// Communication API/ISOBUS/API/bds_isobus_getRxDataboxStatus
///This function reads the current status of one ISOBUS receive databox.
///
///=======
/// Remarks:
///=======
///   + With this function the application can check for every instance of the ISOBUS communication stack whether a ISOBUS databox currently contains valid data.
///   + If the reading of the data is performed outside of a RX callback function then it should be enclosed with the functions BDS_SYS_GET_LOCK_COMMON and BDS_SYS_RELEASE_LOCK_COMMON to ensure data consistency.
///   + This function has to be used to check whether cyclic messages have been received within a defined time interval.
///   + An error state will be automatically reset if the next message has been received correctly.
///   + Instead of polling the RX databox status, the application can also be informed about successfully received data via the RX callback function.
///   + But for the detection of receive timeouts of cyclic PGNs the databox status needs to be polled with this function.
///   + The |GVL_isobus| is given for usage of defines.
///
///
///----------
/// FFI:
///----------
///This API can be used in trusted partitions only. See Freedom from Interference (FFI) concept for more details.
///
///
///==================================================================		  			===================================================================================================
///Return value    								  									Description
///==================================================================		  			===================================================================================================
///16#0000:BDS_ISOBUS_BOXSTATUS_NONE_DU16												Message databox is not yet initialized.
///16#0100:BDS_ISOBUS_BOXSTATUS_INIT_DU16												Message databox is initialized.
///16#0200:BDS_ISOBUS_BOXSTATUS_VALID_DU16												The data within the receive message databox are valid. All data received successfully.
///16#0201:BDS_ISOBUS_BOXSTATUS_VAL_OVFL_DU16											The data within the receive message databox are valid, but incomplete. A buffer overflow occurs (received DM1/2 msg was to long).
///16#0301:BDS_ISOBUS_BOXSTATUS_INV_SEQNBR_DU16										Databox data are invalid, wrong sequence nbr received.
///16#0302:BDS_ISOBUS_BOXSTATUS_INV_ABORT_DU16											Databox data are invalid, rx/tx transfer aborted.
///16#0303:BDS_ISOBUS_BOXSTATUS_INV_TIMEOUT_DU16										Databox data are invalid, timeout occurs.
///16#0304:BDS_ISOBUS_BOXSTATUS_INV_OVFL_DU16											Databox data are invalid, overflow error.
///16#0310:BDS_ISOBUS_BOXSTATUS_INV_PGN_ERR_DU16										Databox data are invalid, different PGN found in RTS and DPO messages.
///16#0311:BDS_ISOBUS_BOXSTATUS_INV_DPO_ERR_DU16										Databox data are invalid, CTS and DPO messages inconsistency.
///16#0500:BDS_ISOBUS_BOXSTATUS_BAM_RX_DU16											Receiving of a BAM message is in progress.
///16#0501:BDS_ISOBUS_BOXSTATUS_CMDT_RX_DU16											Receiving of a CMDT message is in progress.
///16#0700:BDS_ISOBUS_BOXSTATUS_UNPACK_DU16											Unpacking of received DM1/2 BAM is in progress.
///16#0800:BDS_ISOBUS_BOXSTATUS_ETP_RX_DU16											Receiving of an ETP message is in progress.
///
///==================================================================		   			===================================================================================================
///
///=======
///Code Example:
///=======
///============================================================================
///
///VAR_GLOBAL
///
///    (*global data buffer for isobus Rx message*)
///
///    msgRx2Data_au8: ARRAY[1..8] OF USINT;
///
///END_VAR
///
///PROGRAM Isobus_prg
///
///VAR
///
///    len1_u32:UDINT;
///
///    Flag_u8:USINT:=0;
///
///    retval_u16: UINT;
///
///    APPL_ISOBUS_INSTANCES_DU16: USINT:=10;
///
///    isobus_appInst_as:ARRAY[1..10] OF bds_isobus_appInst_ts;
///
///    ISOBUS_RX_BOXES_DU8: USINT:= 5;(* no of rx databoxes*)
///
///    isobus_rxMsg_as: ARRAY[1..5] OF bds_isobus_rxMsg_ts; (*allocate memory for isobus rx databoxes*)
///
///END_VAR
///
///(*call the api once*)
///
///IF(Flag_u8=0)THEN
///    
///    (*registers 10 isobus instances via the below api or by configuring it in easyConfig*)
///
///    bds_isobus_registerInstances(ADR(isobus_appInst_as), APPL_ISOBUS_INSTANCES_DU16);
///    
///    (*register isobus rx message boxes for instance 1*)
///
///    bds_isobus_registerRxDataboxes(1,ADR(isobus_rxMsg_as),ISOBUS_RX_BOXES_DU8);
///    
///    (*initalize rx databox messages for databox 1 of instance 1 with pgn 16#7789*)
///
///    bds_isobus_initRxDatabox(1, 1, 16#7789, 16#04, 2000, 6000, 8,ADR(gvl.msgRx2Data_au8),ADR(Rxcallback));
///    
///    (*define the controller application name, required for address claiming*)
///
///    bds_isobus_setCaName(1,16#00,16#02,16#00,16#01,16#81,16#01,16#01,16#33,BDS_ISOBUS_OWN_SN_DU32);
///    
///    (*define the initial source address and the CAN channel for the CA instance 1*)
///
///    bds_isobus_setCaAddr(1,BDS_CAN_3_D,16#10);
///    
///    (*initialize and start isobus communication for all instances on this CAN channel*)
///
///    bds_isobus_initComm(bds_can_Chnl_te.BDS_CAN_3_D, 50);
///    
///    Flag_u8:=1;
///    
///END_IF
///
///(*check for valid data in a isobus receive databox. Call the Api in cyclic task*)
///
///retval_u16:=bds_isobus_getRxDataboxStatus(1,1, ADR(len1_u32));
///
///
///FUNCTION Rxcallback
///
///VAR
///
///    len_u32:UDINT;
///
///    databox_status_u16: UINT;
///
///END_VAR
///
///(*call the API in callback*)
///
///(*check for valid data in a isobus receive databox.*)
///
///databox_status_u16:=bds_isobus_getRxDataboxStatus(1,1, ADR(len_u32));
///============================================================================
{attribute 'external_name' := 'cmp_rts_bds_isobus_getRxDataboxStatus'}
FUNCTION bds_isobus_getRxDataboxStatus : UINT
VAR_INPUT
	///ISOBUS instance number. This number identifies one instance of the ISOBUS stack.
	///
	///Value range: 1..n
	///n is the number of ISOBUS instances configured by easyConfig. 
	instanceNum_u8: USINT;
	///Number of a ISOBUS receive databox.
	///
	///Value range: 1..n
	///n is the number of receive databoxes configured by easyConfig or alternatively with function |bds_isobus_registerRxDataboxes|
	boxNum_u16: UINT;
	///Pointer to a variable in which the message length [nbr bytes] of the actual received message can be written. If the message length is not required (e.g. PGNs with a fix defined length), then a Null pointer can be given.
	///
	///Exception: If this databox is initialized with the function |bds_isobus_initDiagnostic| for receiving DTCs, then the returned message length is the number of received DTCs.
	msgLen_pu32: POINTER TO UDINT;
END_VAR

END_FUNCTION

// Communication API/ISOBUS/API/bds_isobus_getStatus
///This function reads the current status of an instance of the ISOBUS communication stack.
///
///=======
/// Remarks:
///=======
///   + This function can be called at any time for every instance of the ISOBUS communication stack.
///   + The normal running state of the ISOBUS communication stack is BDS_ISOBUS_CASTATUS_ADDR_CLAIMED_DU16.
///   + In all other main states no messages will be sent.
///   + The return value consists of a main status (high byte) and an independent substatus (low byte).
///   + The |GVL_isobus| is given for usage of defines.
///
///----------
/// FFI:
///----------
///This API can be used in trusted partitions only. See Freedom from Interference (FFI) concept for more details.
///
///==================================================================		  			===================================================================================================
///Return value    								  									Description
///==================================================================		  			===================================================================================================
///Main states:
///16#0000: BDS_ISOBUS_CASTATUS_NONE_DU16												Controller application is not yet initialized, or invalid function parameter.
///16#0100:BDS_ISOBUS_CASTATUS_INIT_DU16												Controller application is initialized.
///16#0200:BDS_ISOBUS_CASTATUS_WAIT_CLAIM_DU16											Controller application waits for answers during an address claim procedure.
///16#0300:BDS_ISOBUS_CASTATUS_ADDR_CLAIMED_DU16										Controller application could claim an address. Message traffic was started.  This is the normal operation state.
///16#0400:BDS_ISOBUS_CASTATUS_CANNOT_CLAIM_DU16										Controller application could not claim an address. There was an address conflict with another controller application. The message traffic will not be started.
///16#FF00: BDS_ISOBUS_CASTATUS_MASK_DU16												This bit mask can be used for the selection of the main status.
///Sub states:																			The sub states may be set in addition to the main states.
///16#0001:BDS_ISOBUS_SUBSTATUS_TIMEOUT_DU16											The ISOBUS communication stack could not handle all ISOBUS messages within one cycle.
///																					   + Possible reasons:
///																						   + The maximum execution time, which is defined with isobus_initComm, is to small.
///																						   + The execution time of one or more callback functions is to high.
///																					   + Remark: This status will be stored until it was read with this function. Afterwards it will be reset automatically.
///16#0002:BDS_ISOBUS_SUBSTATUS_RXOVFL_DU16											There was an overflow of the CAN RX buffer. RX messages may be lost. This error can lead to further protocol errors.
///																					   + Possible reasons:
///																						   + The CAN RX buffer is to small and should be increased.
///																						   + The maximum allowed execution time of the isobus stack is to small and should be increased.
///																					   + Remark: This status will be stored until it was read with this function. Afterwards it will be reset automatically.
///16#0010:BDS_ISOBUS_SUBSTATUS_STOP_BC_DM13_DU16										The DM13 service (Stop Start Broadcast) is active for this controller application. In this status all cyclic broadcast TX messages will be suspended.
///																					   + Possible reasons:	
///																						   + A DM13 message with Stop Broadcast command was received.
///																						   + This status can be quit by receiving a Start Broadcast command.
///
///==================================================================		   			===================================================================================================
///
///=======
///Code Example:
///=======
///============================================================================
///
///PROGRAM appl_Task_1
///
///VAR
///
///	isobusStatus_u16: UINT := 16#00;
///
///END_VAR
///
///
///(* check the isobus communication status of instance 1 *)
///
///isobusStatus_u16 := bds_isobus_getStatus(1);
///
///IF ( BDS_ISOBUS_CASTATUS_ADDR_CLAIMED_DU16 = (isobusStatus_u16 AND BDS_ISOBUS_CASTATUS_MASK_DU16) ) THEN
///
///	(* the address claiming was successful and the ISOBUS communication is running *)
///
///END_IF
///
///============================================================================
{attribute 'external_name' := 'cmp_rts_bds_isobus_getStatus'}
FUNCTION bds_isobus_getStatus : UINT
VAR_INPUT
	///ISOBUS instance number. This number identifies one instance of the ISOBUS stack.
	///
	///Value range: 1..n
	///n is the number of ISOBUS instances configured by easyConfig. 
	instanceNum_u8: USINT;
END_VAR

END_FUNCTION

// I/O API/IN legacy/API/bds_in_sent_disable
///Disables the specified SENT channel.
///
///=======
/// Remarks:
///=======
///   + The disable function of a SENT channel can be used to disable a sensor there are send invalid data.
///
///
///----------
/// FFI:
///----------
///This API can be used in trusted partitions only. See Freedom from Interference (FFI) concept for more details.
///
///==================================================================		  			===================================================================================================
///Return value    								  									Description
///==================================================================		  			===================================================================================================
///0																					No error
///1																					Invalid parameter
///
///==================================================================		   			===================================================================================================
///
///=======
///Code Example:
///=======
///============================================================================
///
///PROGRAM appl_10ms_task
///   VAR
///   
///   END_VAR
///
///  bds_in_sent_disable(bds_in_sent_signal_te.K57);
///  
///END
///
///
///============================================================================
{attribute 'external_name' := 'cmp_rts_bds_in_sent_disable'}
FUNCTION bds_in_sent_disable : USINT
VAR_INPUT
	///The signal name that is assigned to the respective pin configured as SENT input
	signal_e: UINT;
END_VAR

END_FUNCTION

// I/O API/IN legacy/API/bds_in_sent_enable
///Enables the specified SENT channel. 
///
///=======
/// Remarks:
///=======
///   + During startup the BSW enables all SENT inputs, therefore this function needs to be called only if the sent input had been disabled.
///   + The function can be used to re-enable the sent input if disabled.
///
///
///----------
/// FFI:
///----------
///This API can be used in trusted partitions only. See Freedom from Interference (FFI) concept for more details.
///
///==================================================================		  			===================================================================================================
///Return value    								  									Description
///==================================================================		  			===================================================================================================
///0																					No error
///1																					Invalid parameter
///
///==================================================================		   			===================================================================================================
///
///=======
///Code Example:
///=======
///============================================================================
///
///PROGRAM appl_10ms_task
///
///   VAR
///   
///   END_VAR
/// 
///  bds_in_sent_enable(bds_in_sent_signal_te.K57);
///  
///END
///
///============================================================================
{attribute 'external_name' := 'cmp_rts_bds_in_sent_enable'}
FUNCTION bds_in_sent_enable : USINT
VAR_INPUT
	///The signal name that is assigned to the respective pin configured as SENT input
	signal_e: UINT;
END_VAR

END_FUNCTION

// Communication API/ISOBUS/API/bds_isobus_registerErrClrCbk
///This function registers callback functions for DM11 and DM3 respectively for the particular instance.
///
///=======
/// Remarks:
///=======
///   + Received DM3/DM11 automatically clear the isobus failures within the DSM module. The callback can be used to perform additional actions. 
///   + The name of the registered function can be chosen by the user.
///   + If callback is required for only one type of error, other callback function parameter must be passed as NULL.
///   + The |GVL_isobus| is given for usage of defines.
///
///----------
/// FFI:
///----------
///This API can be used in trusted partitions only. See Freedom from Interference (FFI) concept for more details.
///
///==================================================================		  			===================================================================================================
///Return value    								  									Description
///==================================================================		  			===================================================================================================
///None.																				-
///
///==================================================================		   			===================================================================================================
///=======
///Code Example:
///=======
///============================================================================
///
///This Api should be called only once in application.
///
///PROGRAM Isobus_prg
///
///VAR
///    Flag_u8:USINT:=0;    
///
///END_VAR
///
///(*call the api once*)
///
///IF(Flag_u8=0)THEN
///    
///    (* optionally define some ECU information of the controller application for the PGNs HW-ID and SW-ID: *)
///
///    bds_isobus_setCaInfo(2,16#0,ADR(EcuType_as8),ADR(EcuManu_as8),ADR(ApplTask_as8));
///        
///    (*define the controller application name, required for address claiming*)
///
///    bds_isobus_setCaName(1,16#00,16#02,16#00,16#01,16#81,16#01,16#01,16#33,BDS_ISOBUS_OWN_SN_DU32);
///    
///    (*define the initial source address and the CAN channel for the CA instance 1*)
///
///    bds_isobus_setCaAddr(1,BDS_CAN_3_D,16#10);
///    
///    (*initialize and start isobus communication for all instances on this CAN channel*)
///
///    bds_isobus_initComm(bds_can_Chnl_te.BDS_CAN_3_D, 50);
///
///    (*optionally register callback functions for DM3 and DM11*)
///
///    bds_isobus_registerErrClrCbk(2, ADR(isobusDM11Callback), ADR(isobusDM3Callback));
///    
///    Flag_u8:=1;
///    
///END_IF
///
///FUNCTION isobusDM11Callback
///
///VAR
///
///    data_u8: USINT := 16#11;
///
///END_VAR
///
///(*this function will be called when a request PGN DM11 is received*)
///
///bds_can_sendData(2, 16#D11, 1, 1, ADR(data_u8));
///
///FUNCTION isobusDM3Callback
///
///VAR
///
///    data1_u8: USINT := 16#3;
///
///END_VAR
///
///(*this function will be called when a request PGN DM3 is received*)
///
///bds_can_sendData(2, 16#D3, 1, 1, ADR(data1_u8));
///
///============================================================================
{attribute 'external_name' := 'cmp_rts_bds_isobus_registerErrClrCbk'}
FUNCTION bds_isobus_registerErrClrCbk : BOOL
VAR_INPUT
	///ISOBUS instance number. This number identifies one instance of the ISOBUS stack.
	///
	///Value range: 1..n
	///n is the number of ISOBUS instances configured by easyConfig. 
	instanceNum_u8: USINT;
	///Pointer to a callback function to application when DM11 is received.
	DM11func_pf: POINTER TO BOOL;
	///Pointer to a callback function to application when DM3 is received.
	DM3func_pf: POINTER TO BOOL;
END_VAR

END_FUNCTION

// Communication API/ISOBUS/API/bds_isobus_registerTxDataboxes
///This function registers memory for isobus transmit databoxes and therefore defines the maximal number of usable ISOBUS transmit databoxes per instance.
///
///=======
/// Remarks:
///=======
///   + This function must be called once during the configuration of the ISOBUS communication stack before |bds_isobus_initComm|.
///   + After the execution of this function, each isobus transmit databox has to be initialized with |bds_isobus_initTxDatabox| before using.
///   + The DM1/DM2 failure handling, which will be initialized with the function |bds_isobus_initFailureList|, requires 2 additional transmit databoxes.
///   + The |GVL_isobus| is given for usage of defines.
///   + This function should be called only once in the application.
///   
///----------
/// NOTICE:
///----------
///
///This API-function can be used alternatively to the ISOBUS configuration with easyConfig. If this function is used, then the number of ISOBUS TX databoxes is to be configured to 0 in easyConfig.
///
///----------
/// FFI:
///----------
///This API can be used in trusted partitions only. See Freedom from Interference (FFI) concept for more details.
///
///==================================================================		  			===================================================================================================
///Return value    								  									Description
///==================================================================		  			===================================================================================================
///0: BDS_ISOBUS_RC_NO_ERRORS_DU16														Function was executed without errors.
///1: BDS_ISOBUS_RC_INVALID_ADDR_DU16													Address to data array is Invalid.
///8: BDS_ISOBUS_RC_OVERLAP_ADDR_DU16													Address overlaps with an already existing buffer.
///22: BDS_ISOBUS_RC_CFG_NOTALLOWED_DU16												Function must be called before |bds_isobus_initComm|, but it was called afterwards.
///80: BDS_ISOBUS_RC_INV_INST_NUM_DU16													Invalid instance number.
///
///==================================================================		   			===================================================================================================
///
///=======
///Code Example:
///=======
///============================================================================
///
///This Api should be called only once in application.
///
///PROGRAM Isobus_prg
///
///VAR
///
///    Flag_u8:USINT:=0;
///
///    retval_u16: UINT;
///
///    APPL_ISOBUS_INSTANCES_DU16: USINT:=10;
///
///    isobus_appInst_as:ARRAY[1..10] OF bds_isobus_appInst_ts;
///
///    ISOBUS_TX_BOXES_DU8: USINT:= 9; (* no of tx databoxes*)
///
///    isobus_txMsg_as: ARRAY[1..9] OF bds_isobus_txMsg_ts; (*allocate memory for isobus tx databoxes*)   
///
///END_VAR
///
///(*call the api once*)
///
///IF(Flag_u8=0)THEN
///    
///    (*registers 10 isobus instances*)
///
///    bds_isobus_registerInstances(ADR(isobus_appInst_as), APPL_ISOBUS_INSTANCES_DU16);
///    
///    (*register isobus tx message boxes for instance 1*)
///
///    retval_u16:=bds_isobus_registerTxDataboxes(1,ADR(isobus_txMsg_as),ISOBUS_TX_BOXES_DU8);
///
///    Flag_u8:=1;
///    
///END_IF
///
///
///============================================================================
{attribute 'external_name' := 'cmp_rts_bds_isobus_registerTxDataboxes'}
FUNCTION bds_isobus_registerTxDataboxes : UINT
VAR_INPUT
	///ISOBUS instance number. This number identifies one instance of the ISOBUS stack.
	///
	///Value range: 1..n
	///n is the number of ISOBUS instances configured by easyConfig. 
	instanceNum_u8: USINT;
	///Pointer to an array of data type bds_isobus_txMsg_ts.
	///
	///Note:
	///The buffer will be managed by the BSW. The application has only to declare the buffer (memory space).
	///It is necessary to declare the buffer array as a global variable! 
	mem_pas: POINTER TO bds_isobus_txMsg_ts;
	///Size of the array above, which corresponds to the number of usable isobus transmit databoxes.
	num_u16: UINT;
END_VAR

END_FUNCTION

// Communication API/ISOBUS/API/bds_isobus_initTxDatabox
///This function initializes a ISOBUS transmit databox. The ISOBUS messages can be sent only with ISOBUS transmit databoxes.
///
///=======
/// Remarks:
///=======
///   + This function must be called during the configuration of the ISOBUS communication stack once for each ISOBUS transmit message.
///   + Before the TX databoxes can be initialized with this function, the required number of transmit databoxes has to be configured first with easyConfig tool or alternatively with function |bds_isobus_registerTxDataboxes|.
///   + Each ISOBUS TX databox requires an own data array or a data structure. The pointer to this data field is required for the initialization of a ISOBUS transmit databox. The transmitted data will be taken from this data field.
///   + The data array for the transmitted data may have a length of more than 8 bytes (see parameter description below).
///   + The execution time of the callback function should be short to be able to meet the time conditions within the ISOBUS stack. 
///   + If the same CAN bus is also used for further communication, ensure that the CAN IDs are uniquely assigned.
///   + The meaning of this function is similar to the system function |bds_can_initTxDatabox|.
///   + The |GVL_isobus| is given for usage of defines.
///
///----------
/// FFI:
///----------
///This API can be used in trusted partitions only. See Freedom from Interference (FFI) concept for more details.
///
///==================================================================		  			===================================================================================================
///Return value    								  									Description
///==================================================================		  			===================================================================================================
///0: BDS_ISOBUS_RC_NO_ERRORS_DU16														Function was executed without errors.
///2: BDS_ISOBUS_RC_INV_DATABOX_DU16													Invalid databox number.
///3: BDS_ISOBUS_RC_INV_PGN_DU16														Invalid parameter group number (PGN).
///6: BDS_ISOBUS_RC_INV_DATA_LEN_DU16													Invalid data length.
///7: BDS_ISOBUS_RC_INV_DATA_PTR_DU16													Invalid address pointer.
///10: BDS_ISOBUS_RC_INV_CYCLE_DU16													Invalid cycle time.
///11: BDS_ISOBUS_RC_INV_OFFSET_DU16													Invalid offset time.
///12: BDS_ISOBUS_RC_INV_PRIO_DU16														Invalid priority.
///21: BDS_ISOBUS_RC_PGN_PRIO_EXIST_DU16												Another message box with the same PGN and priority is already defined.
///80: BDS_ISOBUS_RC_INV_INST_NUM_DU16													Invalid instance number.
///
///==================================================================		   			===================================================================================================
///
///=======
///Code Example:
///=======
///============================================================================
///
///This Api should be called only once in application.
///
///VAR_GLOBAL
///
///    (*global data buffer for isobus Tx message*)
///
///    msgTx2Data_au8: ARRAY[1..8] OF USINT:=[16#A,2,3,4,5,6,7,8];
///
///END_VAR
///
///PROGRAM Isobus_prg
///
///VAR
///
///    Flag_u8:USINT:=0;
///
///    retval_u16: UINT;
///
///    APPL_ISOBUS_INSTANCES_DU16: USINT:=10;
///
///    isobus_appInst_as:ARRAY[1..10] OF bds_isobus_appInst_ts;
///
///    ISOBUS_TX_BOXES_DU8: USINT:= 9; (* no of tx databoxes*)
///
///    isobus_txMsg_as: ARRAY[1..9] OF bds_isobus_txMsg_ts; (*allocate memory for isobus tx databoxes*)
///
///END_VAR
///
///(*call the api once*)
///
///IF(Flag_u8=0)THEN
///    
///    (*registers 10 isobus instances via the below api or by configuring it in easyConfig*)
///
///    bds_isobus_registerInstances(ADR(isobus_appInst_as), APPL_ISOBUS_INSTANCES_DU16);
///    
///    (*register isobus tx message boxes for instance 1 via the below api or by configuring it in easyConfig*)
///
///    bds_isobus_registerTxDataboxes(1,ADR(isobus_txMsg_as),ISOBUS_TX_BOXES_DU8);
///    
///    (*initalize tx databox messages for databox 3 of instance 1 with pgn 16#1122 in cycle time of 10ms*)
///
///    retval_u16:= bds_isobus_initTxDatabox(1, 3, 16#1122, 6, 10,0, 8,ADR(gvl.msgTx2Data_au8), ADR(Txcallback));
///    
///    (*define the controller application name, required for address claiming*)
///
///    bds_isobus_setCaName(1,16#00,16#02,16#00,16#01,16#81,16#01,16#01,16#33,BDS_ISOBUS_OWN_SN_DU32);
///    
///    (*define the initial source address and the CAN channel for the CA instance 1*)
///
///    bds_isobus_setCaAddr(1,BDS_CAN_3_D,16#10);
///    
///    (*initialize and start isobus communication for all instances on this CAN channel*)
///
///    bds_isobus_initComm(bds_can_Chnl_te.BDS_CAN_3_D, 50);
///    
///    Flag_u8:=1;
///    
///END_IF
///
///(*The data msgTx2Data_au8 to be sent via isobus tx data box 3 can be updated here*)
///
///FUNCTION Txcallback
///
///VAR
///
///END_VAR
///
///IF(gvl.msgTx2Data_au8[1]=16#A) THEN
///
///    gvl.msgTx2Data_au8[3]:=16#C;
///
///END_IF
///============================================================================
{attribute 'external_name' := 'cmp_rts_bds_isobus_initTxDatabox'}
FUNCTION bds_isobus_initTxDatabox : UINT
VAR_INPUT
	///ISOBUS instance number. This number identifies one instance of the ISOBUS stack.
	///
	///Value range: 1..n
	///n is the number of ISOBUS instances configured by easyConfig. 
	instanceNum_u8: USINT;
	///Number of a ISOBUS transmit databox.
	///
	///Value range: 1..n
	///n is the number of transmit databoxes configured by easyConfig or alternatively with function |bds_isobus_registerTxDataboxes|. 
	boxNum_u16: UINT;
	///Parameter group number (PGN) of the message to be sent with this databox.
	///
	///Value range: 0..16#3FFFF (18 bit) 
	///
	///The lowest byte of the PGN contains for:
	///PDU1 format:  the destination address
	///PDU2 format:  the PDU extension
	pgn_u32: UDINT;
	///ISOBUS priority of the message to be sent.
	///
	///Value range: 0..7  (6 = default value according ISOBUS specification) 
	prio_u8: USINT;
	///This time (in ms) controls the cyclic transmission of the ISOBUS message from this ISOBUS databox. The cycle time of a TX message must be greater or equal than the cycle time (= 10ms) of the ISOBUS communication stack. The messages can be only sent with integral multiples of the ISOBUS stack cycle time.
	///
	///With a cycle time = 0 the message will be not sent cyclic. In this case the application may control the sending with the function bds_isobus_sendDatabox().
	///
	///Value range: 10..65000 [ms] or 0 = no cyclic transmission. 
	cycle_u16: UINT;
	///The first transmission cycle of a cyclic ISOBUS message can be shortened by this offset time (in ms). This can be used to prevent CAN bus overload, if several messages have to be sent with the same cycle time. With an offset = 0 the first message will be sent after the cycle time.
	///
	///This parameter is not applicable for cycle_u16 = 0.
	///
	///Value range: 0.. (cycle_u16 - 1) [ms]   
	offset_u16: UINT;
	///Size of the data array/structure below. A ISOBUS message may consist of several single CAN messages, if the number of data bytes is more than 8.
	///
	///Value range: 1..117440512
	lenMax_u32: UDINT;
	///Pointer to a data array or a data structure, from which the data are taken for transmission. The size of this array/structure has to be given within the previous parameter (lenMax_u32).
	///
	///It is neccessary to declare the buffer array/structure as a global variable!
	data_pau8: POINTER TO USINT;
	///Pointer to a callback function of data type UDINT which is called before a new message will be sent. The execution time of the callback function should be short to be able to meet the time conditions within the ISOBUS stack. 
	///The return value of the callback function defines the number of data bytes to which the application may reduce the actual size of the TX message. The return value ISOBUS_BYTES_ALL_DU32 (= 16#FFFFFFFF) sends the message with the whole length as defined within the TX databox.
	///
	///Function must be coded within the application program.
	///Optional a NULL pointer can be assigned to disable the callback function.
	func_pf: POINTER TO UDINT;
END_VAR

END_FUNCTION

// Communication API/ISOBUS/API/bds_isobus_sendDatabox
///This function sends a message from a ISOBUS transmit databox.
///
///=======
/// Remarks:
///=======
///   + This function can be used for sending messages, for which no cycle time is defined.
///   + But this function can also be used for an additional sending of cyclic messages.
///   + The message will be sent not at once, but during the next execution cycle of the ISOBUS communication stack.
///   + The transport protocol of the sending message is dependent on the message definition (PGN, data length) within the transmit databox.
///   + If several messages have to be sent at the same time with a transport protocol like BAM or CMDT, then the messages might be sent delayed. The delay time depends on the occupancy of the corresponding transport protocol handler.
///   + The optionally defined TX callback function will be called right before the message will be sent. In the TX callback function the application may provide actual data.
///   + The ISOBUS cycle time is 10ms.
///   + The |GVL_isobus| is given for usage of defines.
///
///----------
/// FFI:
///----------
///This API can be used in trusted partitions only. See Freedom from Interference (FFI) concept for more details.
///
///==================================================================		  			===================================================================================================
///Return value    								  									Description
///==================================================================		  			===================================================================================================
///0: BDS_ISOBUS_RC_NO_ERRORS_DU16														Function was executed without errors.
///2: BDS_ISOBUS_RC_INV_DATABOX_DU16													Invalid databox number.
///30: BDS_ISOBUS_RC_INV_BOX_STATUS_DU16												Invalid databox status. Databox is not yet initialized or sending of this databox is still in progress. 
///80: BDS_ISOBUS_RC_INV_INST_NUM_DU16													Invalid instance number.
///
///==================================================================		   			===================================================================================================
///
///=======
///Code Example:
///=======
///============================================================================
///
///PROGRAM appl_Task_1
///
///  VAR
///
///  END_VAR
///
///
///  (* send the isobus message from transmit databox 2 of instance 1 *)
///
///  bds_isobus_sendDatabox(1, 2);
///  
///============================================================================
{attribute 'external_name' := 'cmp_rts_bds_isobus_sendDatabox'}
FUNCTION bds_isobus_sendDatabox : UINT
VAR_INPUT
	///ISOBUS instance number. This number identifies one instance of the ISOBUS stack.
	///
	///Value range: 1..n
	///n is the number of ISOBUS instances configured by easyConfig. 
	instanceNum_u8: USINT;
	///Number of a ISOBUS transmit databox.
	///
	///Value range: 1..n
	///n is the number of transmit databoxes configured by easyConfig or alternatively with function |bds_isobus_registerTxDataboxes|. 
	boxNum_u16: UINT;
END_VAR

END_FUNCTION

// Communication API/ISOBUS/API/bds_isobus_initFailureList
///This function initializes the DM1 and DM2 failure handling for the own controller application.
///
///=======
/// Remarks:
///=======
///
///   + This function can be called optionally once for the initialization of the ISOBUS DM1 and DM2 failure handling within the own controller application and it must not be called if the DM1 and DM2 messages are not desired for this instance.
///   + This failure handling requires 2 additional transmit databoxes. They have to be taken into account during the configuration with easyConfig. These 2 databoxes MUST NOT be initialized with the function |bds_isobus_initTxDatabox|.
///   + After the initialization of the failure handling the DM1 message will be sent cyclically every second and the DM2 message will be sent only on request.
///   + This function has no impact on the currently stored DM1/DM2 failures within the system error storage.
///   + The sent DM1/DM2 messages are limited to a size of 32 failures. If the system contains more ISOBUS failures then the list will be truncated to this size.
///   + The |GVL_isobus| is given for usage of defines.
///   + This function should be called only once in the application.
///
///----------
/// FFI:
///----------
///This API can be used in trusted partitions only. See Freedom from Interference (FFI) concept for more details.
///   
///==================================================================		  			===================================================================================================
///Return value    								  									Description
///==================================================================		  			===================================================================================================
///0: BDS_ISOBUS_RC_NO_ERRORS_DU16														Function was executed without errors.
///2: BDS_ISOBUS_RC_INV_DATABOX_DU16													Invalid databox number.
///80: BDS_ISOBUS_RC_INV_INST_NUM_DU16													Invalid instance number.
///
///==================================================================		   			===================================================================================================
///
///=======
///Code Example:
///=======
///============================================================================
///
///This Api should be called only once in application.
///
///PROGRAM Isobus_prg
///
///VAR
///
///    Flag_u8:USINT:=0;
///
///    retval_u16: UINT;
///
///    APPL_ISOBUS_INSTANCES_DU16: USINT:=10;
///
///    isobus_appInst_as:ARRAY[1..10] OF bds_isobus_appInst_ts;
///
///    ISOBUS_TX_BOXES_DU8: USINT:= 9; (* no of tx databoxes*)
///
///    isobus_txMsg_as: ARRAY[1..9] OF bds_isobus_txMsg_ts; (*allocate memory for isobus tx databoxes*)
///
///    dtc2_u16: UINT := 16#8C14;
///
///    result_u16: UINT := BDS_DSM_FAULT_PERCENT_100_DU8;
///
///    statusword_u16: UINT;
///
///    timediff_u32: UDINT := 10000;
///
///END_VAR
///
///(*Configure the DTCs in easyConfig*)
///
///(*Reporting the Error(NoDebounce) with 100 percent fault percentage*)
///
///bds_dsm_updateError_DTC(dtc2_u16, result_u16, timediff_u32);
///
///bds_dsm_getDTC_Status(dtc2_u16, ADR(statusword_u16));
///
///(*call the api once*)
///
///IF(Flag_u8=0)THEN
///    
///    (*registers 10 isobus instances via the below api or by configuring it in easyConfig*)
///
///    bds_isobus_registerInstances(ADR(isobus_appInst_as), APPL_ISOBUS_INSTANCES_DU16);
///    
///    (*register isobus tx message boxes for instance 1 via the below api or by configuring it in easyConfig*)
///
///    bds_isobus_registerTxDataboxes(1,ADR(isobus_txMsg_as),ISOBUS_TX_BOXES_DU8);
///    
///    (*init a DM1 / DM2 failure list for instance 1 on the own ECU*)
///
///    retval_u16:=bds_isobus_initFailureList(1, 8,  9, FALSE);
///        
///    (*define the controller application name, required for address claiming*)
///
///    bds_isobus_setCaName(1,16#00,16#02,16#00,16#01,16#81,16#01,16#01,16#33,BDS_ISOBUS_OWN_SN_DU32);
///    
///    (*define the initial source address and the CAN channel for the CA instance 1*)
///
///    bds_isobus_setCaAddr(1,BDS_CAN_3_D,16#10);
///    
///    (*initialize and start isobus communication for all instances on this CAN channel*)
///
///    bds_isobus_initComm(bds_can_Chnl_te.BDS_CAN_3_D, 50);
///    
///    Flag_u8:=1;
///    
///END_IF
///
///
///============================================================================
{attribute 'external_name' := 'cmp_rts_bds_isobus_initFailureList'}
FUNCTION bds_isobus_initFailureList : UINT
VAR_INPUT
	///ISOBUS instance number. This number identifies one instance of the ISOBUS stack.
	///
	///Value range: 1..n
	///n is the number of ISOBUS instances configured by easyConfig. 
	instanceNum_u8: USINT;
	///The number of a ISOBUS transmit databox, which can be exclusively used for sending of the DM1 message. This databox MUST NOT be initialized additionally with the function bds_isobus_initTxDatabox.
	///
	///Value range: 1..n
	///n is the number of transmit databoxes configured by easyConfig or alternatively with function |bds_isobus_registerTxDataboxes|.
	txBoxDM1_u16: UINT;
	///The number of a ISOBUS transmit databox, which can be exclusively used for sending of the DM2 message. This databox MUST NOT be initialized additionally with the function |bds_isobus_initTxDatabox|.
	///
	///Value range: 1..n
	///n is the number of transmit databoxes configured by easyConfig or alternatively with function |bds_isobus_registerTxDataboxes|.
	txBoxDM2_u16: UINT;
	///Format of lamp status (first 2 bytes) in DM1/2 messages.
	///
	///Possible values:
	///   + TRUE = lamp status according J1939
	///   + FALSE = lamp status according ISOBUS
	j1939Format_l: BOOL;
END_VAR

END_FUNCTION

// Communication API/ISOBUS/API/bds_isobus_sendRequestPGN
///This function requests a PGN (parameter group number) from another controller.
///
///=======
/// Remarks:
///=======
///   + This function can be used to request any PGN from another controller application by sending a message with the PGN RequestPGN (16#00EA00).
///   + This function does not require any ISOBUS transmit databox.
///   + If the AddressClaim PGN (16#00EE00) will be requested with a broadcast request, then the own controller application will answer too.
///   + To be able to receive the answer(s) to the PGN request, the application has to define the corresponding receive databox(es). Exception: Some special PGNs, like the AddressClaim, will be evaluated by the ISOBUS communication stack itself.
///   + The |GVL_isobus| is given for usage of defines.
///
///----------
/// FFI:
///----------
///This API can be used in trusted partitions only. See Freedom from Interference (FFI) concept for more details.
///
///==================================================================		  			===================================================================================================
///Return value    								  									Description
///==================================================================		  			===================================================================================================
///0: BDS_ISOBUS_RC_NO_ERRORS_DU16														Function was executed without errors.
///3: BDS_ISOBUS_RC_INV_PGN_DU16														Invalid parameter group number (PGN).
///50: BDS_ISOBUS_RC_INV_ECU_ADDR_DU16													Invalid controller (ECU) address.
///80: BDS_ISOBUS_RC_INV_INST_NUM_DU16													Invalid instance number.
///
///==================================================================		   			===================================================================================================
///
///=======
///Code Example:
///=======
///============================================================================
///
///PROGRAM Isobus_prg
///
///VAR
///
///    Flag_u8:USINT:=0;
///
///    retval_u16: UINT;
///
///END_VAR
///
///(*call the api once*)
///
///IF(Flag_u8=0)THEN
///        
///    (*define the controller application name, required for address claiming*)
///
///    bds_isobus_setCaName(1,16#00,16#02,16#00,16#01,16#81,16#01,16#01,16#33,BDS_ISOBUS_OWN_SN_DU32);
///    
///    (*define the initial source address and the CAN channel for the CA instance 1*)
///
///    bds_isobus_setCaAddr(1,BDS_CAN_3_D,16#10);
///    
///    (*initialize and start isobus communication for all instances on this CAN channel*)
///
///    bds_isobus_initComm(bds_can_Chnl_te.BDS_CAN_3_D, 50);
///    
///    Flag_u8:=1;
///    
///END_IF
///
///(*request the AddressClaim PGN for instance 1 from controller with address 16#54*)
///
///retval_u16 := bds_isobus_sendRequestPGN(1, 16#54, 16#01789);
///  
///============================================================================
{attribute 'external_name' := 'cmp_rts_bds_isobus_sendRequestPGN'}
FUNCTION bds_isobus_sendRequestPGN : UINT
VAR_INPUT
	///ISOBUS instance number. This number identifies one instance of the ISOBUS stack.
	///
	///Value range: 1..n
	///n is the number of ISOBUS instances configured by easyConfig. 
	instanceNum_u8: USINT;
	///Address of this controller application to which the PGN has to be sent.
	///
	///Value range: 0..253, 255 (=all), own address is not allowed  
	destAddr_u8: USINT;
	///The requested Parameter group number (PGN).
	///
	///Value range: 0..16#3FFFF (18 bit)
	pgn_u32: UDINT;
END_VAR

END_FUNCTION

// Communication API/LIN/API/bds_lin_getStatus
///This function gets the status of the particular LIN channel.
///
///=======
/// Remarks:
///=======
///   + The |GVL_lin| is given for usage of defines.
///   + LIN status information:
///
///
///==========================================		  			==========================================		  			================================================
///Value  								  						Define														Meaning
///==========================================		  			==========================================		  			================================================
///1															BDS_LIN_TX_OK_DU8											Successful transmission.
///2															BDS_LIN_TX_BUSY_DU8											Ongoing transmission (Header or Response).
///3															BDS_LIN_TX_HEADER_ERROR_DU8									Erroneous header transmission such as:
///																														   + Mismatch between the send and read back data.
///																														   + Identifier parity error or physical bus error.
///4															BDS_LIN_TX_ERROR_DU8										Erroneous response transmission such as:
///																														   + Mismatch between the send and read back data.
///																														   + Physical bus error.
///5															BDS_LIN_RX_OK_DU8											Reception of correct response.
///6															BDS_LIN_RX_BUSY_DU8											Ongoing reception: at least one response byte has been received, but the checksum byte has not been received.
///7															BDS_LIN_RX_ERROR_DU8										Erroneous response reception such as:
///																														   + Framing error.
///																														   + Overrun error.
///																														   + Checksum error or Short response.
///8															BDS_LIN_RX_NO_RESPONSE_DU8									No response byte has been received so far.
///9															BDS_LIN_OPERATIONAL_DU8										Normal operation, the related LIN channel is just initialized or waked up from the sleep state and no data has been sent.
///10															BDS_LIN_CH_SLEEP_DU8										Sleep mode operation; in this mode wake-up detection from slave nodes is enabled.
///
///==========================================		  			==========================================					================================================
///
///
///----------
/// FFI:
///----------
///This API can be used in trusted partitions only. See Freedom from Interference (FFI) concept for more details.
///
///==================================================================		  			===================================================================================================
///Return value    								  									Description
///==================================================================		  			===================================================================================================
///BDS_LIN_ERR_NO_ERRORS_DU16 (= 0)													Get status was successful.
///BDS_LIN_INVALID_CHNL_DU16(=121)														Invalid channel.
///BDS_LIN_ERR_NULLPOINTER_DU16(=123)													Invalid address (Null pointer).
///
///==================================================================		   			===================================================================================================
///
///=======
///Code Example:
///=======
///============================================================================
///
///(* the Lin Channel will be available in linCanSignals_easyConfig.xml*)
///
///VAR_GLOBAL
///
///	BDS_LIN_CHNL_1_DU8: USINT := 2;
///	
///END_VAR
///
///PROGRAM appl_task_1
///
///VAR
///
///linSts_u8: USINT := 16#00;
///
///END_VAR
///
///
///(* get the status of particular channel *)
///
///bds_lin_getStatus(BDS_LIN_CHNL_1_DU8, ADR(linSts_u8));
///
///  
///============================================================================
{attribute 'external_name' := 'cmp_rts_bds_lin_getStatus'}
FUNCTION bds_lin_getStatus : UINT
VAR_INPUT
	///LIN channel number.
	channel_u8: USINT;
	///Pointer to the status.
	linstatus_pu8: POINTER TO USINT;
END_VAR

END_FUNCTION

// Communication API/LIN/API/bds_lin_gotoSleep
///This function sends a goto-sleep command on the LIN network for a particular channel.
///
///=======
/// Remarks:
///=======
///   + The LIN goto sleep Frame Counter value can be configured in the cloud tool eC. This value specifies the number of LIN sleep frames to be sent before the LIN channel goes to the sleep state.
///   + The range of goto sleep frame counter value is 1 to 5.
///   + The |GVL_lin| is given for usage of defines.
///
///
///----------
/// FFI:
///----------
///This API can be used in trusted partitions only. See Freedom from Interference (FFI) concept for more details.
///
///==================================================================		  			===================================================================================================
///Return value    								  									Description
///==================================================================		  			===================================================================================================
///BDS_LIN_ERR_NO_ERRORS_DU16 (= 0)													LIN goto-sleep was successful or LIN controller is already in the sleep state.
///BDS_LIN_INVALID_CHNL_DU16 (=121)													Invalid channel.
///
///==================================================================		   			===================================================================================================
///
///=======
///Code Example:
///=======
///============================================================================
///
///(* the Lin Channel will be available in linCanSignals_easyConfig.xml*)
///
///VAR_GLOBAL
///
///	BDS_LIN_CHNL_1_DU8: USINT := 2;
///	
///END_VAR
///
///PROGRAM appl_task_1
///
///VAR
///
///END_VAR
///
///
///(* send the sleep command for a particular channel *)
///
///bds_lin_gotoSleep(BDS_LIN_CHNL_1_DU8);
///
///============================================================================
{attribute 'external_name' := 'cmp_rts_bds_lin_gotoSleep'}
FUNCTION bds_lin_gotoSleep : UINT
VAR_INPUT
	///LIN channel number.
	channel_u8: USINT;
END_VAR

END_FUNCTION

// Communication API/LIN/API/bds_lin_receiveSignal
///Signals are part of PDU/message, call to this API would cause the signal data of the PDU/message received on bus to be copied to application defined buffer.
///
///=======
/// Remarks:
///=======
///   + Cloud tool allows import of LDF file. 
///   + Signals referred here are available upon a valid LDF import. 
///   + For an overview of LIN Protocol, please refer to LIN Overview.
///   + For specific details of integration of LIN into application, please refer to LIN Integration into an application.
///   + The parameters of the signal such as Signal ID, length and signal data pointer are passed as parameters to the function. 
///   + Before receiving the signals the corresponding schedule table under which the signals belong to should be set using |bds_lin_setSchedule| .
///   + The |GVL_lin| is given for usage of defines.
///
///----------
/// FFI:
///----------
///This API can be used in trusted partitions only. See Freedom from Interference (FFI) concept for more details.
///
///-----
/// NOTICE:
///-----
///   + The length parameter specifies the no. of bytes of data to be received and it is important to specify exactly the no. of incoming bytes else it would result in length validation failure.
///   + For signals imported from LDF file, the signal type information comes from LDF. This would generally be of static types like USINT, UINT, SINT, INT.  In order to be able to change the length of signal, it requires that the signal is of type UINT8_DYN. Currently, Easy config cloud tool does not support the selection of signal type to UINT8_DYN. So, for all signals imported from LDF, the length parameter in API has to be set to 0.
///   + Signal IDs can be located in the post build configuration file - linCanSignals_easyConfig.xml. 
///   
///==================================================================		  			===================================================================================================
///Return value    								  									Description
///==================================================================		  			===================================================================================================
///BDS_LIN_ERR_NO_ERRORS_DU16 (= 0)													Signal reception successful.
///BDS_LINSIG_ERR_RX_FAIL_DU16(=118)													Reception failure.
///BDS_LINSIG_ERR_RX_NOSERVICE_DU16(=120)												Service not available - PDU inactive.
///BDS_LINSIG_ERR_RX_DATAPTR_DU16(=115)												Invalid data pointer address.
///BDS_LINSIG_ERR_NUM_RX_SIG_DU16(=113)												Invalid Signal ID.
///
///==================================================================		   			===================================================================================================
///
///=======
///Code Example:
///=======
///============================================================================
///
///(* the schedule table entry and the signals present in LDF file and imported via eC will be available in linCanSignals_easyConfig.xml*)
///
///VAR_GLOBAL
///
///	BDS_LIN_CHNL_1_DU8: USINT := 2;
///	
///	ComSignal_LIN_LIN_Power_Out_H: USINT := 10;
///	
///	LinIf_rbr_RUN_HEATER_LinIfChannel_0_LinIfGlobalConfig_0: USINT := 16#03;
///	
///END_VAR
///
///PROGRAM Lin_prg
///
///    Rx_data_au8: USINT;
///	
///    length_au16:UINT:= 0;
///	
///    flag:UINT:=0;
///	
///VAR
///
///(*call the api once*)
///
///IF(flag=0) THEN 
///   
///    (*set the schedule table*)
///
///    bds_lin_setSchedule(BDS_LIN_CHNL_1_DU8,LinIf_rbr_RUN_HEATER_LinIfChannel_0_LinIfGlobalConfig_0);
///	
///    flag:=1;
///	
///END_IF
///
///IF( 0 = bds_lin_receiveSignal(ComSignal_LIN_LIN_Power_Out_H,ADR(Rx_data_au8), length_au16) ) THEN
///
/// (* ok,Data is stored in Rx_data_au8 *)
///
///END_IF
///
///============================================================================
{attribute 'external_name' := 'cmp_rts_bds_lin_receiveSignal'}
FUNCTION bds_lin_receiveSignal : UINT
VAR_INPUT
	///ID of the signal to be received.
	signalId_u16: UINT;
	///Pointer array to location where the received signal data shall be stored.
	signalDataPtr_au8: POINTER TO USINT;
	///No. of bytes of data expected to be received (for dynamic type signal)
	///- 0 , for static signals (imported from LDF,refer NOTICE above).
	length_u16: UINT;
END_VAR

END_FUNCTION

// Communication API/LIN/API/bds_lin_setSchedule
///This function is used to set a particular schedule table for a specific LIN channel.This function is used to set a particular schedule table for a specific LIN channel.
///
///=======
/// Remarks:
///=======
///   + Cloud tool allows import of LDF file.
///   + The Schedule tables present in the LDF file can only be used in the application. Addition of separate schedule table in eC is not supported.
///   + To stop the LIN communication the |bds_lin_setSchedule| should be used with the NULL_SCHEDULE as parameter.
///   + The |GVL_lin| is given for usage of defines.
///
///
///----------
/// FFI:
///----------
///This API can be used in trusted partitions only. See Freedom from Interference (FFI) concept for more details.
///
///==================================================================		  			===================================================================================================
///Return value    								  									Description
///==================================================================		  			===================================================================================================
///BDS_LIN_ERR_NO_ERRORS_DU16 (= 0)													Schedule table request successful.
///BDS_LIN_INVALID_CHNL_DU16(=121u)													Invalid channel.
///BDS_LIN_INVALID_SCHTABLE_NO_DU16(=122u)												Invalid schedule table number.
///
///
///==================================================================		   			===================================================================================================
///
///=======
///Code Example:
///=======
///============================================================================
///
///(* the schedule table entry and the lin channel present in LDF file and imported via eC will be available in linCanSignals_easyConfig.xml*)
///
///VAR_GLOBAL
///
///	BDS_LIN_CHNL_1_DU8: USINT := 2;
///	
///	LinIf_rbr_RUN_HEATER_LinIfChannel_0_LinIfGlobalConfig_0: USINT := 16#03;
///	
///END_VAR
///
///
///PROGRAM Lin_prg
///	
///    flag:UINT:=0;
///	
///VAR
///
///(*call the api once*)
///
///IF(flag=0) THEN 
///   
///    (*set the schedule table*)
///
///    bds_lin_setSchedule(BDS_LIN_CHNL_1_DU8,LinIf_rbr_RUN_HEATER_LinIfChannel_0_LinIfGlobalConfig_0);
///	
///    flag:=1;
///	
///END_IF
///
///
///(* Set the null schedule table to stop the LIN communication *)
///
///bds_lin_setSchedule(BDS_LIN_CHNL_1_DU8, NULL_SCHEDULE);
///
///============================================================================
{attribute 'external_name' := 'cmp_rts_bds_lin_setSchedule'}
FUNCTION bds_lin_setSchedule : UINT
VAR_INPUT
	///LIN channel number.
	channel_u8: USINT;
	///Schedule table number.
	scheduleTblNo_u8: USINT;
END_VAR

END_FUNCTION

// Communication API/LIN/API/bds_lin_sendSignal
///This function is used to transmit message with signal data specified by signal ID on the LIN bus.
///
///Signals are part of PDU , call to this API would cause the PDU to be sent on bus but with the signal contents updated by the signal data pointer.
///
///=======
/// Remarks:
///=======
///   + Cloud tool allows import of LDF file.
///   + Signals referred here are available upon a valid LDF import. 
///   + For an overview of LIN Protocol, please refer to  LIN Overview.
///   + For specific details of integration of LIN into application, please refer to LIN Integration into an application.
///   + The parameters of the signal such as Signal ID, length and signal data pointer are passed as parameters to the function.
///   + Before sending the signals the corresponding schedule table under which the signals belong to should be set using |bds_lin_setSchedule|.
///   + The |GVL_lin| is given for usage of defines.
///
///----------
/// FFI:
///----------
///This API can be used in trusted partitions only. See Freedom from Interference (FFI) concept for more details.
///
///-----
/// NOTICE:
///-----
///   + For signals imported from LDF file, the signal type information comes from LDF. This would generally  be of static types like USINT, UINT, SINT, INT.  In order to be able to change the length of signal, it requires that the signal is of type UINT8_DYN. Presently, Easy config cloud tool does not support the selection of signal type to UINT8_DYN. So, for   all signals imported from LDF, the length parameter in API has to be set to 0.
///   + Signal IDs can be located in the post build configuration file - linCanSignals_easyConfig.xml. 
///   
///==================================================================		  			===================================================================================================
///Return value    								  									Description
///==================================================================		  			===================================================================================================
///BDS_LIN_ERR_NO_ERRORS_DU16 (= 0)													Signal transmission successful.
///BDS_LINSIG_ERR_TX_FAIL_DU16(=117u)													Transmission failure.
///BDS_LINSIG_ERR_TX_NOSERVICE_DU16(=119)												Service not available-PDU inactive.
///BDS_LINSIG_ERR_TX_DATAPTR_DU16(=114)												Invalid data pointer address.
///BDS_LINSIG_ERR_NUM_TX_SIG_DU16(=112)												Invalid Signal ID.
///
///==================================================================		   			===================================================================================================
///
///=======
///Code Example:
///=======
///============================================================================
///
///(* the schedule table entry and the signals  present in LDF file and imported via eC will be available in linCanSignals_easyConfig.xml*)
///
///VAR_GLOBAL
///
///	BDS_LIN_CHNL_1_DU8: USINT := 2;
///	
///	ComSignal_LIN_LIN_CTRL_PWR_H: USINT := 9;
///	
///	LinIf_rbr_RUN_HEATER_LinIfChannel_0_LinIfGlobalConfig_0: USINT := 16#03;
///	
///END_VAR
///
///PROGRAM Lin_prg
///
///    signaldata_au8:USINT:=16#7;
///	
///    length_au16:UINT:= 0;
///	
///    flag:UINT:=0;
///	
///VAR
///
///(*call the api once*)
///
///IF(flag=0) THEN 
///   
///    (*set the schedule table*)
///
///    bds_lin_setSchedule(BDS_LIN_CHNL_1_DU8,LinIf_rbr_RUN_HEATER_LinIfChannel_0_LinIfGlobalConfig_0);
///	
///    flag:=1;
///	
///END_IF
///
///IF( 0 = bds_lin_SendSignal(ComSignal_LIN_LIN_CTRL_PWR_H,ADR(signaldata_au8),length_au16) ) THEN
///
/// (* ok,message is sent on bus with updated signal data *)
///
///END_IF
///
///
///============================================================================
{attribute 'external_name' := 'cmp_rts_bds_lin_sendSignal'}
FUNCTION bds_lin_sendSignal : UINT
VAR_INPUT
	///ID of the signal to be sent.
	signalId_u16: UINT;
	///Pointer array to the signal data to be transmitted.
	signalDataPtr_au8: POINTER TO USINT;
	///-No. of bytes of data to be sent (for dynamic type signal)
	///- 0 , for static signals(imported from LDF, refer NOTICE above).
	length_u16: UINT;
END_VAR

END_FUNCTION

// I/O API/OUT_LEGACY/bds_out_aov_cfg
///Configures the voltage deviation for an analog voltage output.
///
///=======
/// Remarks:
///=======
///   + Maximal allowed deviation between the set point and the actual voltage is 500mV. The signal quality of the PWM must be considered for the deviation value.    
///   + For more information see |bds_out_aov_getStatus|.
///   + This function should be called only once in the application.
///
///----------
/// FFI:
///----------
///This API can be used in trusted partitions . For untrusted partitions use |bds_out_aov_cfg_ffi|. See Freedom from Interference (FFI) concept for more details.
///   
///==================================================================		  			===================================================================================================
///Return value    								  									Description
///==================================================================		  			===================================================================================================
///0																					No error
///1																					Invalid parameter
///
///==================================================================		   			===================================================================================================
///
///=======
///Code Example:
///=======
///============================================================================
///
///PROGRAM PLC_PRG
///
///  VAR
///  
///	Init_flag_u8:USINT:=0;
/// 
///  END_VAR
///  
///IF(Init_flag_u8=0) THEN (*To make api call once in application*)
///
///	(* set a deviation of 100mV for output K62 (e.g. once at start up) *)
///	
///	bds_out_aov_cfg(bds_out_aov_signal_te.K62, 100);
///  
///	Init_flag_u8:=1;
///  
///END_IF
///
///============================================================================
{attribute 'external_name' := 'cmp_rts_bds_out_aov_cfg'}
FUNCTION bds_out_aov_cfg : USINT
VAR_INPUT
	///The connector assigned signal name of the output
	signal_e: UINT;
	///Allowed voltage deviation [mV].Range:
	///   + 0 to 500
	uDeviation_u16: UINT;
END_VAR

END_FUNCTION

// I/O API/OUT_LEGACY/bds_out_aov_getStatus
///Provides status of an analog voltage output.
///
///=======
/// Remarks:
///=======
///   + The status data holds all relevant information of the analog voltage output.
///	   + Part of the status data is also the fault status of every DFC (e.g. stDFC_SCB_u16).
///	   + With the macros (e.g. bds_dsm_DFC_ldf) defined in bds_dsm_api.h , respective bit fields of the fault status can be read.
///
///----------
/// FFI:
///----------
///This API can be used in trusted partitions . For untrusted partitions use |bds_out_aov_getStatus_ffi|. See Freedom from Interference (FFI) concept for more details.
///
///==================================================================		  			===================================================================================================
///Return value    								  									Description
///==================================================================		  			===================================================================================================
///0																					No error
///1																					Invalid parameter
///
///==================================================================		   			===================================================================================================
///
///=======
///Code Example:
///=======
///============================================================================
///
///PROGRAM appl_10ms_task
///
///VAR
///
/// 	stK62_s: bds_out_aov_ts;
///
/// 	ldf_u8: USINT := 16#00;
///
///END_VAR
///
///(* get the status of output K62 *)
///
///bds_out_aov_getStatus(bds_out_aov_signal_te.K62, ADR(stK62_s));
///
///
///(* get last debounced fault *)
///
///ldf_u8 = bds_dsm_DFC_ldf(stK62_s.stDFC_SCB_u16);
///
///============================================================================
{attribute 'external_name' := 'cmp_rts_bds_out_aov_getStatus'}
FUNCTION bds_out_aov_getStatus : USINT
VAR_INPUT
	///The connector assigned signal name of the output.
	signal_e: UINT;
	///Storage address of the data. pointer to |bds_out_aov_ts|
	data_ps: POINTER TO bds_out_aov_ts;
END_VAR

END_FUNCTION

// I/O API/OUT/FFI_API/bds_out_aov_getStatus_ffi
{attribute 'external_name' := 'cmp_rts_bds_out_aov_getStatus_ffi'}
FUNCTION bds_out_aov_getStatus_ffi : USINT
VAR_INPUT
	///The connector assigned signal name of the output.
	signal_e: UINT;
	///Storage address of the data. pointer to |bds_out_aov_ts|
	data_ps: POINTER TO bds_out_aov_ts;
END_VAR

END_FUNCTION

// I/O API/OUT/FFI_API/bds_out_aov_cfg_ffi
{attribute 'external_name' := 'cmp_rts_bds_out_aov_cfg_ffi'}
FUNCTION bds_out_aov_cfg_ffi : USINT
VAR_INPUT
	///The connector assigned signal name of the output
	signal_e: UINT;
	///Allowed voltage deviation [mV].Range:
	///   + 0 to 500
	uDeviation_u16: UINT;
END_VAR

END_FUNCTION

// I/O API/OUT_LEGACY/bds_out_aov_cfgPI
///Sets the gain values for Kp and Ki of a analog voltage output.
///
///=======
/// Remarks:
///=======
///   + The range of Kp is defined as 0..2000 and for Ki as 0..500.
///   + The default values after reset of the ECU are Kp = 100 and Ki = 25.
///   + For more information see |bds_out_aov_getStatus|
///   + The information about definitions and structures can be found in  BODAS API library, bds_rts_ec.xml.
///
///----------
/// FFI:
///----------
///This API can be used in trusted partitions . For untrusted partitions use |bds_out_aov_cfgPI_ffi|. See Freedom from Interference (FFI) concept for more details.
///
///==================================================================		  			===================================================================================================
///Return value    								  									Description
///==================================================================		  			===================================================================================================
///0																					No error
///1																					Invalid parameter
///
///==================================================================		   			===================================================================================================
///
///=======
///Code Example:
///=======
///============================================================================
///
///PROGRAM PLC_PRG
///
///VAR
///
///END_VAR
///
///(* configure the gain values for output K25 *)
///
///bds_out_aov_cfgPI(bds_out_aov_signal_te.K25, 200, 100);
///
///============================================================================
{attribute 'external_name' := 'cmp_rts_bds_out_aov_cfgPI'}
FUNCTION bds_out_aov_cfgPI : USINT
VAR_INPUT
	///The connector assigned signal name of the output. See bds_out_aov_signal_te in bds_rts_ec.xml.
	signal_e: UINT;
	///Kp value
	///   + Range:0..2000
	///   + Default : 100
	kp_u16: UINT;
	///Ki value
	///   + Range:0..500
	///   + Default : 25
	ki_u16: UINT;
END_VAR

END_FUNCTION

// I/O API/OUT/FFI_API/bds_out_aov_cfgPI_ffi
{attribute 'external_name' := 'cmp_rts_bds_out_aov_cfgPI_ffi'}
FUNCTION bds_out_aov_cfgPI_ffi : USINT
VAR_INPUT
	///The connector assigned signal name of the output. See bds_out_aov_signal_te in bds_rts_ec.xml.
	signal_e: UINT;
	///Kp value
	///   + Range:0..2000
	///   + Default : 100
	kp_u16: UINT;
	///Ki value
	///   + Range:0..500
	///   + Default : 25
	ki_u16: UINT;
END_VAR

END_FUNCTION

// I/O API/OUT_LEGACY/bds_out_aov_getVoltage
///Provides  voltage of an analog voltage output.
///
///=======
/// Remarks:
///=======
///   + The voltage range depends on the type.
///	   + AOV: 0 to 12000mV
///	   + PWM: 0 to 33000mV.
///   + The read-back path of the voltage can also be used as analog input if the set point is set to zero. ( see also |bds_out_aov|). Diagnostics capabilities similar to standard inputs is not available. 
///
///----------
/// FFI:
///----------
///This API can be used in trusted partitions . For untrusted partitions use |bds_out_aov_getVoltage_ffi|. See Freedom from Interference (FFI) concept for more details.
///
///------
/// Info:
///------
///
///For the predefined type AOV is also a reconfiguration with the eC tool as analog voltage input or digital input possible.
///
///==================================================================		  			===================================================================================================
///Return value    								  									Description
///==================================================================		  			===================================================================================================
///0																					No error
///1																					Invalid parameter
///2																					Function call was erroneous.
///
///==================================================================		   			===================================================================================================
///
///=======
///Code Example:
///=======
///============================================================================
///
///PROGRAM appl_10ms_task
///
///VAR
///
/// 	uK62_u16: UINT := 16#00;
///
///END_VAR
///
/// 
///
///(* get voltage of output K62 *)
///
///bds_out_aov_getVoltage(bds_out_aov_signal_te.K62, ADR(uK62_u16));
///
///============================================================================
{attribute 'external_name' := 'cmp_rts_bds_out_aov_getVoltage'}
FUNCTION bds_out_aov_getVoltage : USINT
VAR_INPUT
	///The connector assigned signal name of the output.
	signal_e: UINT;
	///Storage address of the value.Range:
	///   + AOV: 0 to 12000mV
	///   + PWM: 0 to 33000mV
	value_pu16: POINTER TO UINT;
END_VAR

END_FUNCTION

// I/O API/OUT_LEGACY/bds_out_aov
///Sets the analog voltage output to a given set point.
///
///=======
/// Remarks:
///=======
///   + The analog voltage has two output types namely PWM and AOV. 
///	   + The set point range of the PWM is 25 to 75% of the battery voltage.
///	   + The set point range of the AOV is 0 to 10000mV.
///	   + If the set point has been set to 0 value then the output can also be used as analog voltage input. (see |bds_out_aov_getVoltage|)
///   + For more information see |bds_out_aov_getStatus| and |bds_out_aov_resetError|.
///
///----------
/// FFI:
///----------
///This API can be used in trusted partitions . For untrusted partitions use |bds_out_aov_ffi|. See Freedom from Interference (FFI) concept for more details.
///
///------
/// Info:
///------
///
///For the output type PWM an external load is mandatory, see Technical Data Sheet (RE-sheet RE95207).
///
///
///==================================================================		  			===================================================================================================
///Return value    								  									Description
///==================================================================		  			===================================================================================================
///0																					No error
///1																					Invalid parameter
///2																					Output is locked
///
///==================================================================		   			===================================================================================================
///
///=======
///Code Example:
///=======
///============================================================================
///
///PROGRAM appl_10ms_task
///
///VAR
///
///END_VAR
///
///(* set a voltage of 50% of Ubat for type PWM *)
///
///bds_out_aov(bds_out_aov_signal_te.K25, 500);
///
///(* set a voltage of 5000mV for type AOV *)
///
///bds_out_aov(bds_out_aov_signal_te.K62, 5000);
///
///============================================================================
{attribute 'external_name' := 'cmp_rts_bds_out_aov'}
FUNCTION bds_out_aov : USINT
VAR_INPUT
	///The connector assigned signal name of the output.
	signal_e: UINT;
	///New set point for PWM [0.1%] respective AOV [mV].Range:
	///   + PWM: 0 and 250 to 750
	///   + AOV: 0 to 10000
	uSet_u16: UINT;
END_VAR

END_FUNCTION

// I/O API/OUT_LEGACY/bds_out_aov_resetError
///Resets an error and unlocks the analog voltage output.
///
///
///==================================================================		  			===================================================================================================
///Return value    								  									Description
///==================================================================		  			===================================================================================================
///0																					No error
///1																					Invalid parameter
///
///==================================================================		   			===================================================================================================
///
///----------
/// FFI:
///----------
///This API can be used in trusted partitions only. See Freedom from Interference (FFI) concept for more details.
///
///=======
///Code Example:
///=======
///============================================================================
///
///PROGRAM appl_10ms_task
///
///VAR
///
///	return_u8: USINT := 16#00;
///
///END_VAR
///
///
///
///(* reset error of output K62 *)
///
///return_u8 = bds_out_aov_resetError(bds_out_aov_signal_te.K62);
///
///
///============================================================================
{attribute 'external_name' := 'cmp_rts_bds_out_aov_resetError'}
FUNCTION bds_out_aov_resetError : USINT
VAR_INPUT
	///The connector assigned signal name of the output.
	signal_e: UINT;
END_VAR

END_FUNCTION

// I/O API/OUT/FFI_API/bds_out_aov_ffi
{attribute 'external_name' := 'cmp_rts_bds_out_aov_ffi'}
FUNCTION bds_out_aov_ffi : USINT
VAR_INPUT
	///The connector assigned signal name of the output.
	signal_e: UINT;
	///New set point for PWM [0.1%] respective AOV [mV].Range:
	///   + PWM: 0 and 250 to 750
	///   + AOV: 0 to 10000
	uSet_u16: UINT;
END_VAR

END_FUNCTION

// I/O API/OUT/FFI_API/bds_out_aov_getVoltage_ffi
{attribute 'external_name' := 'cmp_rts_bds_out_aov_getVoltage_ffi'}
FUNCTION bds_out_aov_getVoltage_ffi : USINT
VAR_INPUT
	///The connector assigned signal name of the output.
	signal_e: UINT;
	///Storage address of the value.Range:
	///   + AOV: 0 to 12000mV
	///   + PWM: 0 to 33000mV
	value_pu16: POINTER TO UINT;
END_VAR

END_FUNCTION

// I/O API/OUT_LEGACY/bds_out_cfgLoadCharacteristic
///Configures the load characteristics for a pair of outputs.
///
///By default the ECU including BODAS-API is designed to drive loads with inductive impedance .
///
///In case the application wants to drive loads with different characteristics e.g. capacitive impedance, the application has to configure the load's characteristics with this function.
///
///=======
/// Remarks:
///=======
///   + Whenever the application sets the load characteristic type to capacitive impedance (load_characteristic_e = CAPACITIVE_LOAD. see parameter below), the following applies:
///	   + Open load detection of the high side is suppressed.
///	   + Short circuit to ground and open load detection of the low side is only performed as long as the output is turned on.
///	   + Short circuit to battery is not detected whenever the outputs are turned off.
///   + The high side output will be driven in proportional mode
///   + The low side output will be driven in digital mode.
///   + If one of the chosen outputs is already used for  configuration of a safout channel or as power supply for the low sides this is indicated with the return value.  See  |bds_safout_cfg| and |bds_out_po_cfgPwrLs|.
///   + This function should be called only once in the application.
///
///----------
/// FFI:
///----------
///This API can be used in trusted partitions . For untrusted partitions use |bds_out_cfgLoadCharacteristic_ffi|. See Freedom from Interference (FFI) concept for more details.
///   
///------
/// Info:
///------
///
///Currently this function supports the transition from default (inductive) to capacitive mode only.
///
///==================================================================		  			===================================================================================================
///Return value    								  									Description
///==================================================================		  			===================================================================================================
///0																					No error
///1																					Invalid parameter
///2																					Proportional output already configured
///3																					Digital output already configured
///
///==================================================================		   			===================================================================================================
///
///=======
///Code Example:
///=======
///============================================================================
///
///PROGRAM PLC_PRG
///
///VAR
///
///	Init_flag_u8:USINT:=0;
///
///END_VAR
///  
///IF(Init_flag_u8=0) THEN (*To make api call once in application*)
///
///	(* configure a proportional and a digital output for configuring the loader characteristic *)
///	
///	bds_out_cfgLoadCharacteristic(bds_out_po_signal_te.K07, bds_out_po_signal_te.K12, 1);
///  
///	Init_flag_u8:=1;
///  
///END_IF
///
///PROGRAM appl_100ms_task
///
///VAR
///
///END_VAR
///
///
///
///(* switch loader lights on *)
///
///bds_out_pod(bds_out_po_signal_te.K07, STD_ACTIVE);
///
///bds_out_do(bds_out_po_signal_te.K12, STD_ACTIVE);
///
///
///
///(* switch loader lights off *)
///
///bds_out_pod(bds_out_po_signal_te.K07, STD_IDLE);
///
///bds_out_do(bds_out_po_signal_te.K12, STD_IDLE);
///
///============================================================================
{attribute 'external_name' := 'cmp_rts_bds_out_cfgLoadCharacteristic'}
FUNCTION bds_out_cfgLoadCharacteristic : USINT
VAR_INPUT
	///The connector assigned signal name of the proportional  high side output.
	signal_po_e: UINT;
	///The connector assigned signal name of the digital low side output.
	signal_do_e: UINT;
	///This parameter has to be set to CAPACITIVE_LOAD if the application wants to run such load. Otherwise no action from the application is needed.
	///   + 0 = INDUCTIVE_LOAD
	///   + 1 = CAPACITIVE_LOAD
	///   
	///NOTE: if "INDUCTIVE_LOAD" is used, the function does not perform any action as this is the default mode. The function returns "a parameter is invalid".
	load_characteristic_e: bds_load_characteristic_te;
END_VAR

END_FUNCTION

// I/O API/OUT/FFI_API/bds_out_cfgLoadCharacteristic_ffi
{attribute 'external_name' := 'cmp_rts_bds_out_cfgLoadCharacteristic_ffi'}
FUNCTION bds_out_cfgLoadCharacteristic_ffi : USINT
VAR_INPUT
	///The connector assigned signal name of the proportional  high side output.
	signal_po_e: UINT;
	///The connector assigned signal name of the digital low side output.
	signal_do_e: UINT;
	///This parameter has to be set to CAPACITIVE_LOAD if the application wants to run such load. Otherwise no action from the application is needed.
	///   + 0 = INDUCTIVE_LOAD
	///   + 1 = CAPACITIVE_LOAD
	///   
	///NOTE: if "INDUCTIVE_LOAD" is used, the function does not perform any action as this is the default mode. The function returns "a parameter is invalid".
	load_characteristic_e: bds_load_characteristic_te;
END_VAR

END_FUNCTION

// I/O API/OUT_LEGACY/bds_out_do_cfgPwrLs
///Configures a proportional high side output as power supply for the low side outputs.
///
///=======
/// Remarks:
///=======
///   + The output is also switched on with the configuration.
///   + If the output is switched off and switched on again with bds_out_do the open load faults of the connected low sides must be reset using |bds_out_po_resetError| or |bds_out_do_resetError| depending on the configuration of the output.
///   + A high side output must be used for the power supply of the low sides because a direct supply on the low side outputs is not permitted, see also Proportional outputs and Digital outputs.
///
///----------
/// FFI:
///----------
///This API can be used in trusted partitions  For untrusted partitions use |bds_out_do_cfgPwrLs_ffi|. See Freedom from Interference (FFI) concept for more details.
///
///------
/// Info:
///------
///
///With this configuration the open load detection is suppressed for the high side output. Therefore the output shall be configured during the start up of the RC, otherwise a fault may be detected depending on the time of configuration.
///
///==================================================================		  			===================================================================================================
///Return value    								  									Description
///==================================================================		  			===================================================================================================
///0																					No error
///1																					A parameter is invalid.
///2																					Function call was erroneous.
///3																					Output is not in use (Disabled)
///4																					Output is disabled.
///5																					output is locked 
///6																					Output is already configured. 
///
///==================================================================		   			===================================================================================================
{attribute 'external_name' := 'cmp_rts_bds_out_do_cfgPwrLs'}
FUNCTION bds_out_do_cfgPwrLs : USINT
VAR_INPUT
	///The connector assigned signal name of the high side output. See bds_out_do_signal_te in bds_rts_ec.xml.
	signal_e: UINT;
END_VAR

END_FUNCTION

// I/O API/OUT/FFI_API/bds_out_do_cfgPwrLs_ffi
{attribute 'external_name' := 'cmp_rts_bds_out_do_cfgPwrLs_ffi'}
FUNCTION bds_out_do_cfgPwrLs_ffi : USINT
VAR_INPUT
	///The connector assigned signal name of the high side output. See bds_out_do_signal_te in bds_rts_ec.xml.
	signal_e: UINT;
END_VAR

END_FUNCTION

// I/O API/OUT_LEGACY/bds_out_do_disable
///Disables unused digital output to avoid the setting of faults.
///
///=======
/// Remarks:
///=======
///   + Prevents the setting of open load faults at an unused output.
///   + The output should be disabled during start up.
///   + This function should be called only once in the application.
///
///----------
/// FFI:
///----------
///This API can be used in trusted partitions . For untrusted partitions use |bds_out_do_disable_ffi|. See Freedom from Interference (FFI) concept for more details.
///
///------
/// Attention:
///------
///
///If an output is  disabled, faults are not longer detected and also the control of the output is suppressed
///
///==================================================================		  			===================================================================================================
///Return value    								  									Description
///==================================================================		  			===================================================================================================
///0																					No error
///1																					Invalid parameter
///2																					Output is already configured as safout, output can't be disabled
///
///==================================================================		   			===================================================================================================
///
///=======
///Code Example:
///=======
///============================================================================
///
///PROGRAM PLC_PRG
///
///VAR
///
///	Init_flag_u8:USINT:=0;
///
///END_VAR
///  
///IF(Init_flag_u8=0) THEN (*To make api call once in application*)
///
///	(* disable output K87 *)
///	
///	bds_out_do_disable(bds_out_do_signal_te.K87, STD_ON);
///	
///	Init_flag_u8:=1;
///  
///END_IF
///
///============================================================================
{attribute 'external_name' := 'cmp_rts_bds_out_do_disable'}
FUNCTION bds_out_do_disable : USINT
VAR_INPUT
	///The connector assigned signal name of the output.
	signal_e: UINT;
	///The states are
	///   + STD_OFF - Enable the output (default)
	///   + STD_ON   - Disable the output
	state_u8: USINT;
END_VAR

END_FUNCTION

// I/O API/OUT/FFI_API/bds_out_do_disable_ffi
{attribute 'external_name' := 'cmp_rts_bds_out_do_disable_ffi'}
FUNCTION bds_out_do_disable_ffi : USINT
VAR_INPUT
	///The connector assigned signal name of the output.
	signal_e: UINT;
	///The states are
	///   + STD_OFF - Enable the output (default)
	///   + STD_ON   - Disable the output
	state_u8: USINT;
END_VAR

END_FUNCTION

// Communication API/LIN/API/bds_lin_wakeUp
///This function sends a wake-up request on the LIN network for a particular channel and wake-up the bus if it is in the sleep state.
///
///=======
/// Remarks:
///=======
///   + After the call of wake-up function, it is required to call the |bds_lin_setSchedule| function to start the communication again.
///   + The |GVL_lin| is given for usage of defines.
///
///----------
/// FFI:
///----------
///This API can be used in trusted partitions only. See Freedom from Interference (FFI) concept for more details.
///
///
///==================================================================		  			===================================================================================================
///Return value    								  									Description
///==================================================================		  			===================================================================================================
///BDS_LIN_ERR_NO_ERRORS_DU16 (= 0)													LIN wake-up was successful or the controller is not in sleep state.
///BDS_LIN_INVALID_CHNL_DU16(=121u)													Invalid channel.
///
///==================================================================		   			===================================================================================================
///
///=======
///Code Example:
///=======
///============================================================================
///
///(* the schedule table entry and the lin channel present in LDF file and imported via eC will be available in linCanSignals_easyConfig.xml*)
///
///VAR_GLOBAL
///
///	BDS_LIN_CHNL_1_DU8: USINT := 2;
///	
///	LinIf_rbr_RUN_HEATER_LinIfChannel_0_LinIfGlobalConfig_0: USINT := 16#03;
///	
///END_VAR
///
///PROGRAM Lin_prg
///	
///    flag:UINT:=0;
///	
///VAR
///
///(* send the wake-up command for a particular channel *)
///
///bds_lin_wakeUp(BDS_LIN_CHNL_1_DU8);
///
///
///
///(* After the call of wake-up , the set schedule function should be called to restart the communication *)
///
///(* Set the required schedule table entry *)
///
///(* the schedule table entry present in LDF file and imported via eC will be available in linCanSignals_easyConfig.xml*)
///
///(*call the api once*)
///
///IF(flag=0) THEN 
///   
///    (*set the schedule table*)
///
///    bds_lin_setSchedule(BDS_LIN_CHNL_1_DU8,LinIf_rbr_RUN_HEATER_LinIfChannel_0_LinIfGlobalConfig_0);
///	
///    flag:=1;
///	
///END_IF
///
///============================================================================
{attribute 'external_name' := 'cmp_rts_bds_lin_wakeUp'}
FUNCTION bds_lin_wakeUp : UINT
VAR_INPUT
	///LIN channel number.
	channel_u8: USINT;
END_VAR

END_FUNCTION

// I/O API/OUT_LEGACY/bds_out_do_disableTstPls
///Disables test pulses for a dedicated digital output to avoid having test pulses for error detection on that output.
///
///=======
/// Remarks:
///=======
///   + Test pulses are enabled by default.
///   + For some application this test pulses disturb the wanted functionality of the output for example if you want to use it for power supply.
///   + The test pulses can be deactivated for High Power Outputs only.
///   + This function should be called only once in the application.
/// 
///----------
/// FFI:
///----------
///This API can be used in trusted partitions . For untrusted partitions use |bds_out_do_disableTstPls_ffi|. See Freedom from Interference (FFI) concept for more details.
///  
///------
/// Attention:
///------
///
///If test pulses are disabled, for an output then the fault detection and healing is limited.
///
///==================================================================		  			===================================================================================================
///Return value    								  									Description
///==================================================================		  			===================================================================================================
///0																					No error
///1																					Signal is out of range.
///2																					State Command out of range.
///3																					Output is configured as safout, Test pulse can't be disabled
///
///==================================================================		   			===================================================================================================
///
///=======
///Code Example:
///=======
///============================================================================
///
///PROGRAM PLC_PRG
///
///VAR
///
///	Init_flag_u8:USINT:=0;
///
///END_VAR
///  
///IF(Init_flag_u8=0) THEN (*To make api call once in application*)
///
///	(* disable test pulses for output K13 *)
///	
///	bds_out_do_disableTstPls(bds_out_do_signal_te.K13, STD_ON);
///	
///	Init_flag_u8:=1;
///  
///END_IF
///
///============================================================================
{attribute 'external_name' := 'cmp_rts_bds_out_do_disableTstPls'}
FUNCTION bds_out_do_disableTstPls : USINT
VAR_INPUT
	///The connector assigned signal name of the output.
	signal_e: UINT;
	///The states are
	///   + STD_OFF -  Enables the test pulses (default
	///   + STD_ON   - Disable the test pulses
	state_u8: USINT;
END_VAR

END_FUNCTION

// I/O API/OUT/FFI_API/bds_out_do_disableTstPls_ffi
{attribute 'external_name' := 'cmp_rts_bds_out_do_disableTstPls_ffi'}
FUNCTION bds_out_do_disableTstPls_ffi : USINT
VAR_INPUT
	///The connector assigned signal name of the output.
	signal_e: UINT;
	///The states are
	///   + STD_OFF -  Enables the test pulses (default
	///   + STD_ON   - Disable the test pulses
	state_u8: USINT;
END_VAR

END_FUNCTION

// I/O API/OUT_LEGACY/bds_out_do_getCurrent
///Provides current on a digital output.
///
///=======
/// Remarks:
///=======
///   + The current measurement and corresponding current sensing is just possible for the high power outputs.
///   + The threshold for the over current detection is 6000mA and therefore also the measurement range is defined from 0 to 6000mA.
///   + For more information see |bds_out_do_getStatus|.
///
///
///----------
/// FFI:
///----------
///This API can be used in trusted partitions . For untrusted partitions use |bds_out_do_getCurrent_ffi|. See Freedom from Interference (FFI) concept for more details.
///
///==================================================================		  			===================================================================================================
///Return value    								  									Description
///==================================================================		  			===================================================================================================
///0																					No error
///1																					A parameter is invalid.
///2																					Current measurement unit not available for the output
///
///==================================================================		   			===================================================================================================
///
///=======
///Code Example:
///=======
///============================================================================
///
///PROGRAM appl_10ms_task
///
///VAR
///
///	iK12_u16: UINT := 16#00;
///
///END_VAR
///
///
///
///(* get the current of output K12 *)
///
///bds_out_do_getCurrent(bds_out_do_signal_te.K12, ADR(iK12_u16));
///
///
///============================================================================
{attribute 'external_name' := 'cmp_rts_bds_out_do_getCurrent'}
FUNCTION bds_out_do_getCurrent : USINT
VAR_INPUT
	///The connector assigned signal name of the output.
	signal_e: UINT;
	///Storage address of the value.
	///
	///   + Range:0 to 60000 [mA]
	value_pu16: POINTER TO UINT;
END_VAR

END_FUNCTION

// I/O API/OUT/FFI_API/bds_out_do_getCurrent_ffi
{attribute 'external_name' := 'cmp_rts_bds_out_do_getCurrent_ffi'}
FUNCTION bds_out_do_getCurrent_ffi : USINT
VAR_INPUT
	///The connector assigned signal name of the output.
	signal_e: UINT;
	///Storage address of the value.
	///
	///   + Range:0 to 60000 [mA]
	value_pu16: POINTER TO UINT;
END_VAR

END_FUNCTION

// System API/DSM/API/bds_dsm_getErrorsJ1939
///This function is used to get all DTCs with the specified status configured for J1939 only.
///
///=======
/// Remarks:
///=======
///    + The |GVL_dsm| is given for usage of defines.
///	+ Suspect Parameter Number (SPN), Failure Mode Identifier (FMI) and Lamp States can be configured in easyConfig.
///
///----------
/// FFI:
///----------
///This API can be used in trusted partitions only. See Freedom from Interference (FFI) concept for more details.
///
///-----
/// NOTICE:
///-----
///	+ On a maximum, 32 different DFES entries are possible 
///	+ This function can return maximum 32 entries.
///	+ SPN or FMI should be non zero to be visible in J1939.
///	
///==================================================================		  			===================================================================================================
///Return value    								  									Description
///==================================================================		  			===================================================================================================
///16#0000: BDS_DSM_NO_ERROR_DU16														Update Number of Error is Successful .
///16#0004: BDS_DSM_INVALID_PTR_DU16													Invalid Pointer.
///16#0005: BDS_DSM_STATE_ERROR_DU16													Invalid State.
///16#000A: BDS_DSM_WRONG_BUFFERSIZE_DU16												Buffersize is invalid.
///16#000B:BDS_DSM_NO_DTC_AVAILABLE_DU16												No more DTC is available.
///
///==================================================================		   			===================================================================================================
///
///
///=======
///Code Example:
///=======
///============================================================================
///
///PROGRAM DSM
///
///VAR
///
///	mask_s : UINT := BDS_DSM_SET_ACTIVE_ERROR_MASK_DU16;
///
///	startFromBegin_l: BOOL := TRUE;
///
///	maxNum_u16:USINT := 32;
///
///	error_count_u16: UINT;
///
///	dfc_active_s: ARRAY [1..32] OF bds_dsm_J1939_info_ts;
///
///	status_u16: UINT;
///
///END_VAR
///
///
///(*Get the number of error starting from the begin*)
///
///status_u16 := bds_dsm_getErrorsJ1939(ACTIVE_ERRORS,ADR(dfc_active_s),startFromBegin_L,maxNum_u16,ADR(error_count_u16));
///
///IF status_u16 = BDS_DSM_NO_ERROR_DU16 THEN
///
///	(*Number of Errors has been read successfully*)
///
///END_IF
///
///
///============================================================================
///
{attribute 'external_name' := 'cmp_rts_bds_dsm_getErrorsJ1939'}
FUNCTION bds_dsm_getErrorsJ1939 : UINT
VAR_INPUT
	///The kind of error status can be specified in detail by means of this mask.
	///    + ACTIVE_ERRORS(0)                      - Fault is Active.
	///    + PREVIOUSLY_ACTIVE_ERRORS(1) - Fault was Previously Active.
	state_e: bds_dsm_state_te;
	///pointer to a variable where the DTC data is returned.
	DTC_buffer_ts: POINTER TO bds_dsm_J1939_info_ts;
	///
	///    + TRUE: Query is started from the beginning of DFES.
	///    + FALSE: Query is continued with the next index where the last query was finished.
	startFromBegin_l: BOOL;
	///maximal number of errors/DTCs which can be returned.
	bds_buffersize_u8: USINT;
	///pointer to a variable where the number of errors/DTCs are returned.
	bds_count_DTC_u8: POINTER TO USINT;
END_VAR

END_FUNCTION

